(* Logix 5000 project; controller TFF vendor 1 type 14 code 107 rev 33.11; software revision 33.04; part 37 of 38 *)
(* tags used below, declared in another part *)
   Config : Configuration;   // Index Array used in configuration routines
   result : DINT[2];
   SCL : SCALE;   // Scale Instruction
   AI101Alarm : ALIAS FOR AlarmAnalog[16];
   AI104Alarm : ALIAS FOR AlarmAnalog[17];
   ControlLoop_TIC101Alarm : ALIAS FOR AlarmDeviation[7];
   FlowPath : FlowPath[64];   // Flow Path Array
   LI101 : ALIAS FOR AnalogPoint[44];
   LI101Alarm : ALIAS FOR AlarmAnalog[44];
   Options : Options;   // Options List
   PI601Alarm : ALIAS FOR AlarmAnalog[21];
   PipeAnimation : PipeAnimation;   // HMI Pipe Animation Array
   Rack_ACT350_WI101_200L : IO_Station;   // Status of ACT350 200L
   Rack_ACT350_WI101_500L : IO_Station;   // Status of ACT350 500L
   Tank : TankManagement;   // Tank Management
   TCU101Alarm : ALIAS FOR AlarmAnalog[18];
   TCU101DF : ALIAS FOR DigitalPoint[30];
   TI101Alarm : ALIAS FOR AlarmAnalog[13];
   WI101 : ALIAS FOR AnalogPoint[15];
   WI101Alarm : ALIAS FOR AlarmAnalog[15];
(* Process, continued *)

ROUTINE TankManagement   (* ladder *)
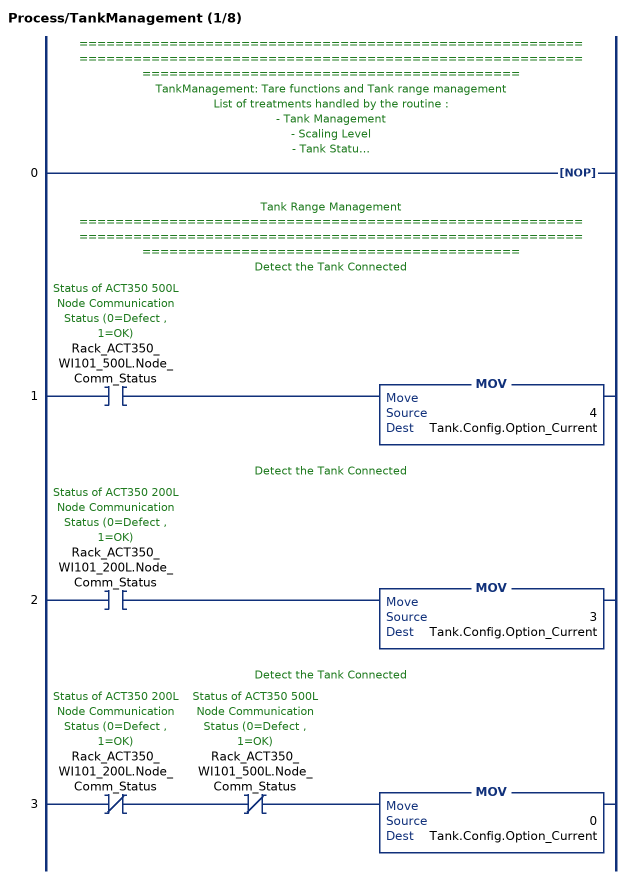
   // ==========================================================================================================================================================
   //                                                                                                                                 TankManagement: Tare functions and Tank range management
   //                                                     List of treatments handled by the routine :
   //                                                          - Tank Management
   //                                                          - Scaling Level
   //                                                          - Tank Status
   //                                                     -----------------------------------------------------------------------------------------------------------------------------------------------------
   //                                                     History
   // 		2019-DEC-24 - Merck - Q. Spindler - Initial version for Candidate Release 1.00.00.00.a
   // ==========================================================================================================================================================
   0: NOP();
   // Tank Range Management
   // ==========================================================================================================================================================
   // Detect the Tank Connected
   1: XIC(Rack_ACT350_WI101_500L.Node_Comm_Status)MOV(4,Tank.Config.Option_Current);
   // Detect the Tank Connected
   2: XIC(Rack_ACT350_WI101_200L.Node_Comm_Status)MOV(3,Tank.Config.Option_Current);
   // Detect the Tank Connected
   3: XIO(Rack_ACT350_WI101_200L.Node_Comm_Status)XIO(Rack_ACT350_WI101_500L.Node_Comm_Status)MOV(0,Tank.Config.Option_Current);
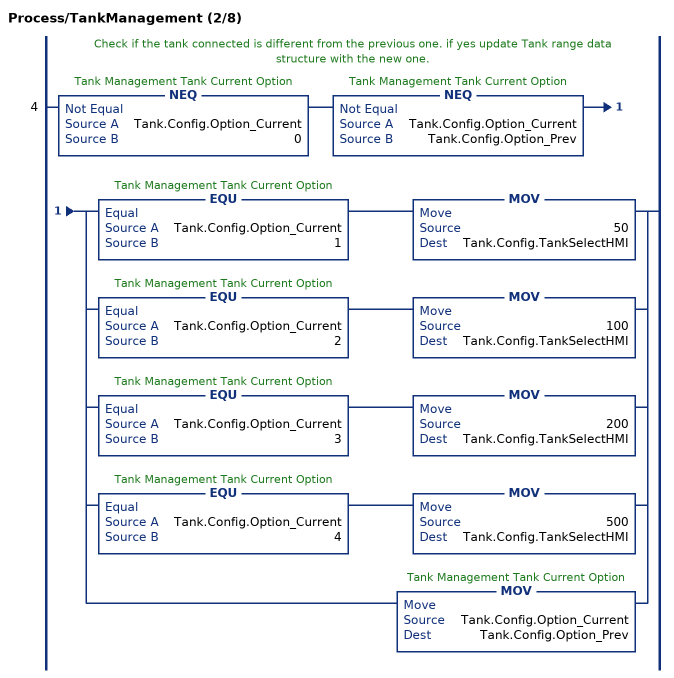
   // Check if the tank connected is different from the previous one. if yes update Tank range data structure with the new one.
   4: NEQ(Tank.Config.Option_Current,0)NEQ(Tank.Config.Option_Current,Tank.Config.Option_Prev)[[EQU(Tank.Config.Option_Current,1) MOV(50,Tank.Config.TankSelectHMI) ,EQU(Tank.Config.Option_Current,2) MOV(100,Tank.Config.TankSelectHMI) ,EQU(Tank.Config.Option_Current,3) MOV(200,Tank.Config.TankSelectHMI) ,EQU(Tank.Config.Option_Current,4) MOV(500,Tank.Config.TankSelectHMI) ] ,MOV(Tank.Config.Option_Current,Tank.Config.Option_Prev) ];
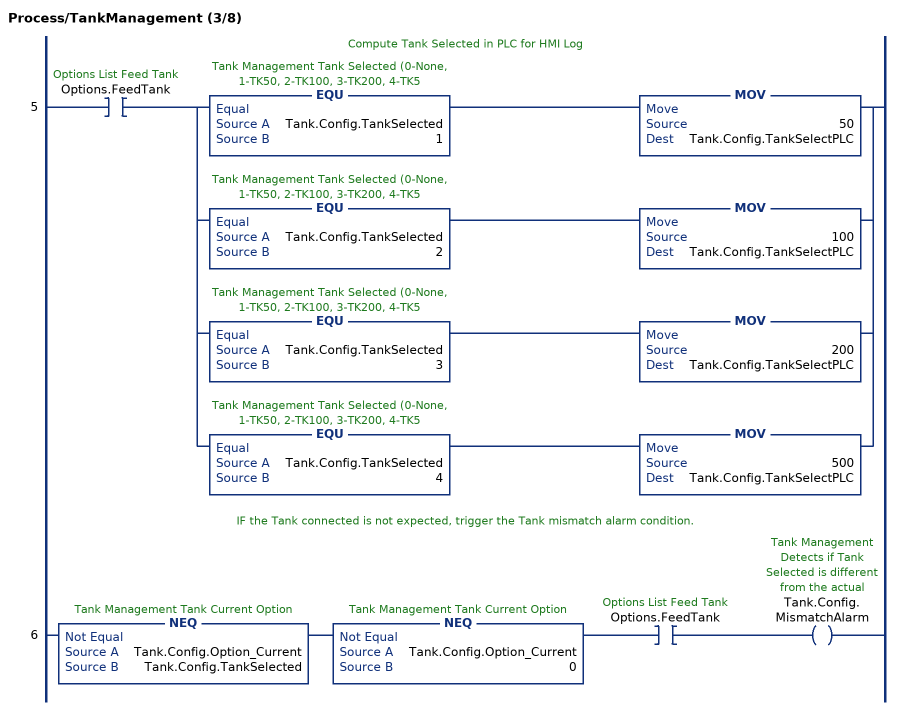
   // Compute Tank Selected in PLC for HMI Log
   5: XIC(Options.FeedTank)[EQU(Tank.Config.TankSelected,1) MOV(50,Tank.Config.TankSelectPLC) ,EQU(Tank.Config.TankSelected,2) MOV(100,Tank.Config.TankSelectPLC) ,EQU(Tank.Config.TankSelected,3) MOV(200,Tank.Config.TankSelectPLC) ,EQU(Tank.Config.TankSelected,4) MOV(500,Tank.Config.TankSelectPLC) ];
   // IF the Tank connected is not expected, trigger the Tank mismatch alarm condition.
   6: NEQ(Tank.Config.Option_Current,Tank.Config.TankSelected)NEQ(Tank.Config.Option_Current,0)XIC(Options.FeedTank)OTE(Tank.Config.MismatchAlarm);
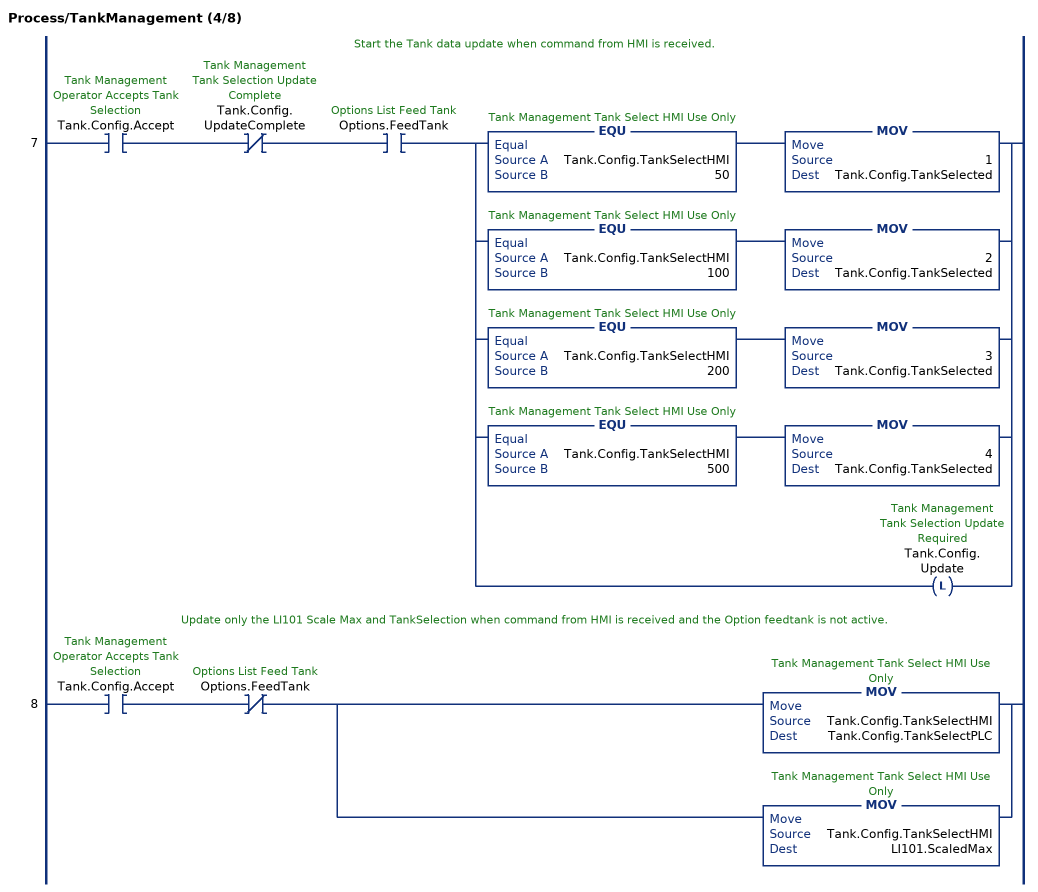
   // Start the Tank data update when command from HMI is received.
   7: XIC(Tank.Config.Accept)XIO(Tank.Config.UpdateComplete)XIC(Options.FeedTank)[[EQU(Tank.Config.TankSelectHMI,50) MOV(1,Tank.Config.TankSelected) ,EQU(Tank.Config.TankSelectHMI,100) MOV(2,Tank.Config.TankSelected) ,EQU(Tank.Config.TankSelectHMI,200) MOV(3,Tank.Config.TankSelected) ,EQU(Tank.Config.TankSelectHMI,500) MOV(4,Tank.Config.TankSelected) ] ,OTL(Tank.Config.Update) ];
   // Update only the LI101 Scale Max and TankSelection when command from HMI is received and the Option feedtank is not active.
   8: XIC(Tank.Config.Accept)XIO(Options.FeedTank)[MOV(Tank.Config.TankSelectHMI,Tank.Config.TankSelectPLC) ,MOV(Tank.Config.TankSelectHMI,LI101.ScaledMax) ];
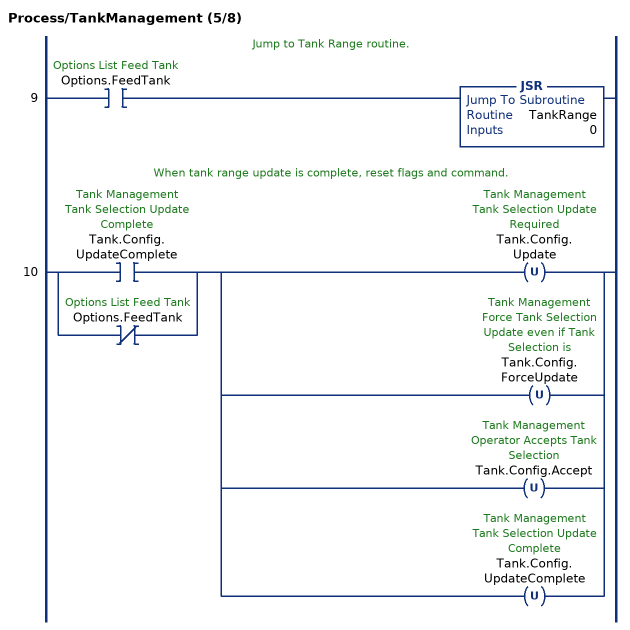
   // Jump to Tank Range routine.
   9: XIC(Options.FeedTank)JSR(TankRange,0);
   // When tank range update is complete, reset flags and command.
   10: [XIC(Tank.Config.UpdateComplete) ,XIO(Options.FeedTank) ][OTU(Tank.Config.Update) ,OTU(Tank.Config.ForceUpdate) ,OTU(Tank.Config.Accept) ,OTU(Tank.Config.UpdateComplete) ];
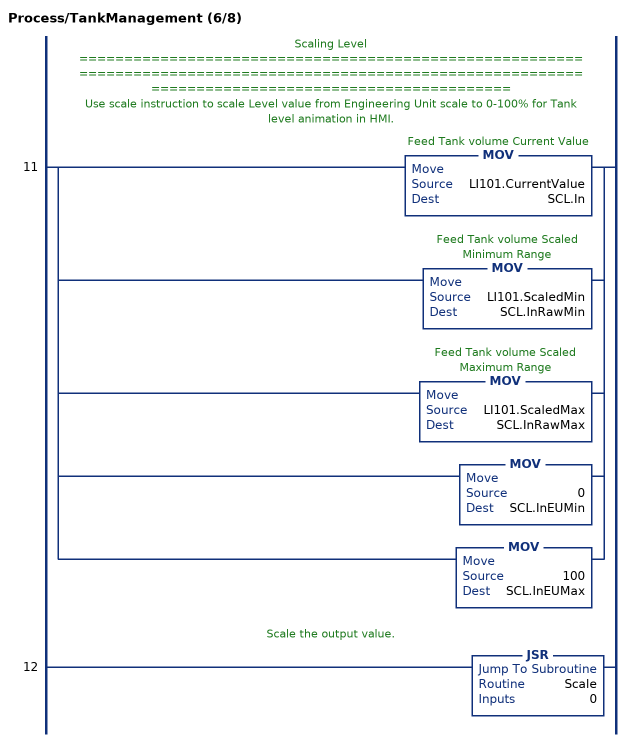
   // Scaling Level
   // ========================================================================================================================================================
   // Use scale instruction to scale Level value from Engineering Unit scale to 0-100% for Tank level animation in HMI.
   11: [MOV(LI101.CurrentValue,SCL.In) ,MOV(LI101.ScaledMin,SCL.InRawMin) ,MOV(LI101.ScaledMax,SCL.InRawMax) ,MOV(0,SCL.InEUMin) ,MOV(100,SCL.InEUMax) ];
   // Scale the output value.
   12: JSR(Scale,0);
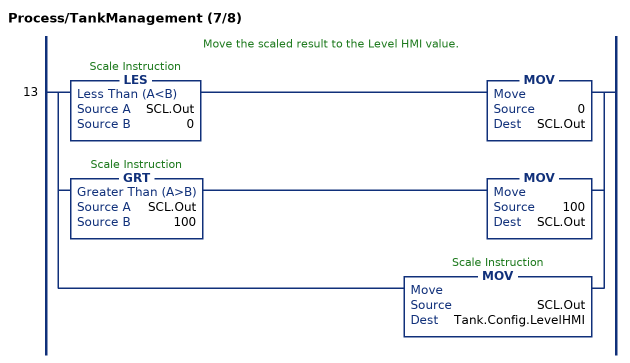
   // Move the scaled result to the Level HMI value.
   13: [LES(SCL.Out,0) MOV(0,SCL.Out) ,GRT(SCL.Out,100) MOV(100,SCL.Out) ,MOV(SCL.Out,Tank.Config.LevelHMI) ];
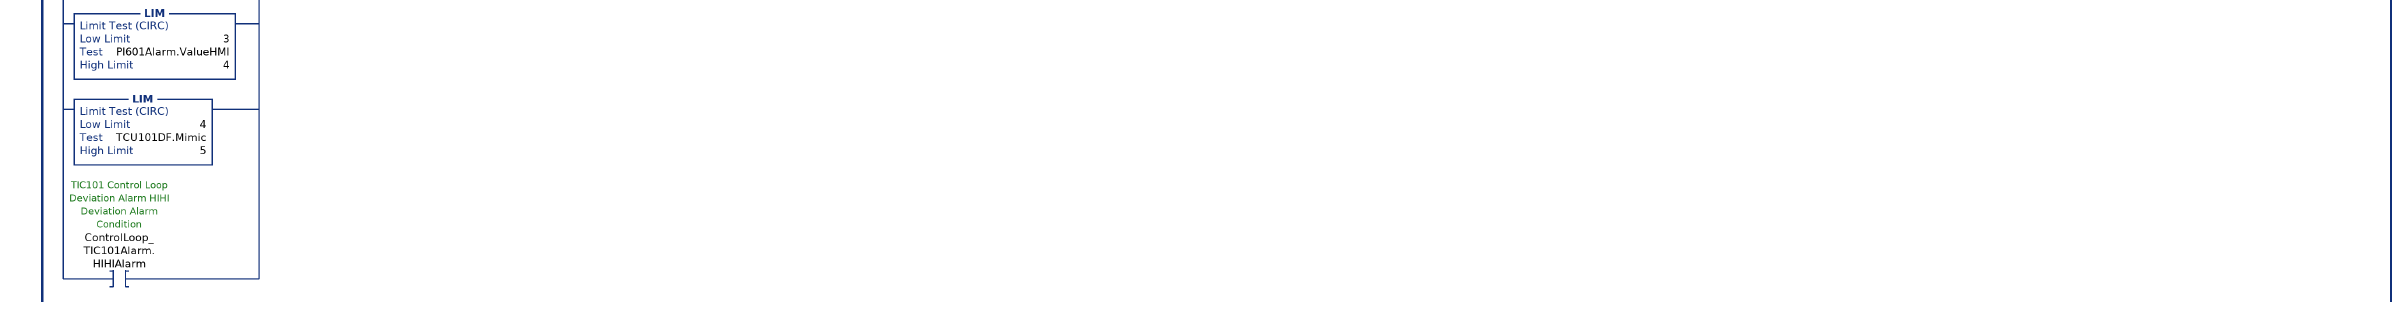
   // Tank Status
   // ==========================================================================================================================================================
   // TankAlarmStatus : 0 = No Alarm & No Flowpath Valid
   // TankAlarmStatus : 1 = No Alarm & Flowpath Valid
   // TankAlarmStatus : 2 = Tank in Non-Critical Alarm
   // TankAlarmStatus : 3 = Tank in Critical Alarm
   14: [XIO(PipeAnimation.PipeStatP1[23]) XIO(PipeAnimation.PipeStatP2[10]) LES(WI101Alarm.ValueHMI,1) LES(LI101Alarm.ValueHMI,1) LES(TI101Alarm.ValueHMI,1) LES(TCU101Alarm.ValueHMI,1) LES(AI101Alarm.ValueHMI,1) LES(AI104Alarm.ValueHMI,1) LES(PI601Alarm.ValueHMI,1) LES(TCU101DF.Mimic,2) XIO(ControlLoop_TIC101Alarm.HIAlarm) XIO(ControlLoop_TIC101Alarm.HIHIAlarm) MOV(0,Tank.Config.AlarmStatus) ,[XIC(PipeAnimation.PipeStatP1[23]) ,XIC(PipeAnimation.PipeStatP2[10]) ] LES(WI101Alarm.ValueHMI,1) LES(LI101Alarm.ValueHMI,1) LES(TI101Alarm.ValueHMI,1) LES(TCU101Alarm.ValueHMI,1) LES(AI101Alarm.ValueHMI,1) LES(AI104Alarm.ValueHMI,1) LES(PI601Alarm.ValueHMI,1) LES(TCU101DF.Mimic,2) XIO(ControlLoop_TIC101Alarm.HIAlarm) XIO(ControlLoop_TIC101Alarm.HIHIAlarm) MOV(1,Tank.Config.AlarmStatus) ,[LIM(1,WI101Alarm.ValueHMI,2) ,LIM(1,LI101Alarm.ValueHMI,2) ,LIM(1,TI101Alarm.ValueHMI,2) ,LIM(1,TCU101Alarm.ValueHMI,2) ,LIM(1,AI101Alarm.ValueHMI,2) ,LIM(1,AI104Alarm.ValueHMI,2) ,LIM(1,PI601Alarm.ValueHMI,2) ,LIM(2,TCU101DF.Mimic,3) ,XIC(ControlLoop_TIC101Alarm.HIAlarm) XIO(ControlLoop_TIC101Alarm.HIHIAlarm) ] MOV(2,Tank.Config.AlarmStatus) ,[LIM(3,WI101Alarm.ValueHMI,4) ,LIM(3,LI101Alarm.ValueHMI,4) ,LIM(3,TI101Alarm.ValueHMI,4) ,LIM(3,TCU101Alarm.ValueHMI,4) ,LIM(3,AI101Alarm.ValueHMI,4) ,LIM(3,AI104Alarm.ValueHMI,4) ,LIM(3,PI601Alarm.ValueHMI,4) ,LIM(4,TCU101DF.Mimic,5) ,XIC(ControlLoop_TIC101Alarm.HIHIAlarm) ] MOV(3,Tank.Config.AlarmStatus) ];
END_ROUTINE

ROUTINE TankRange   (* ladder *)
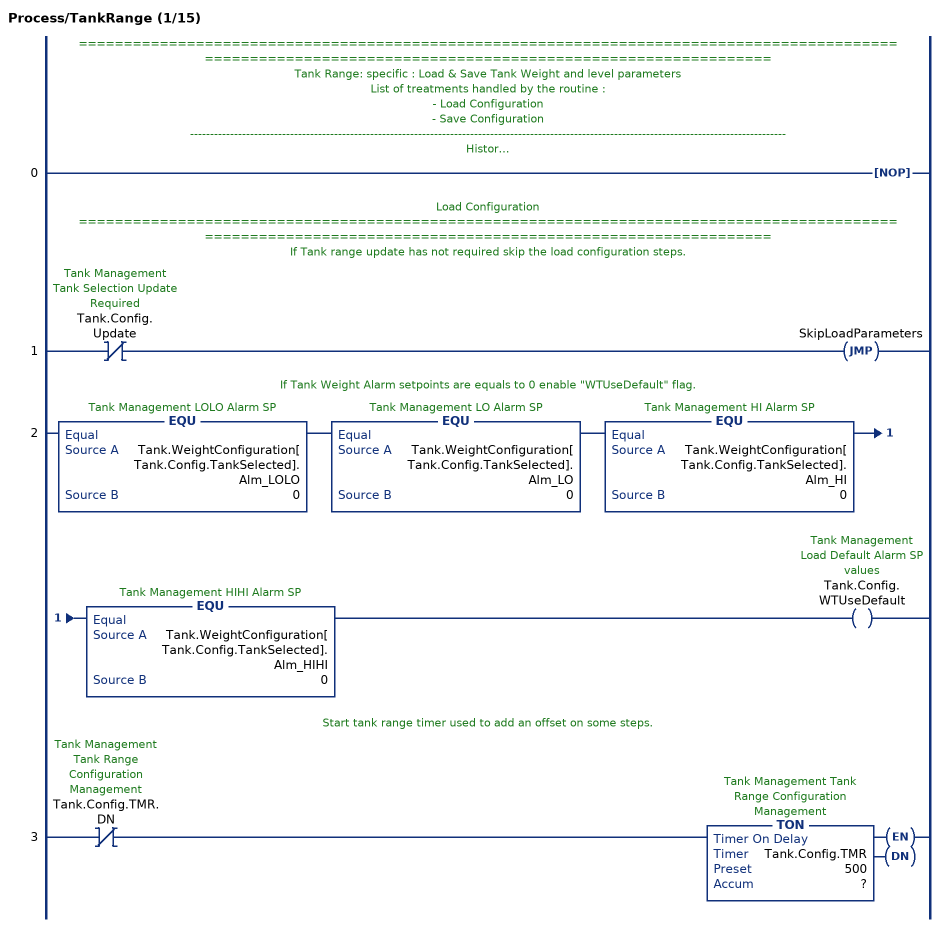
   // ==========================================================================================================================================================
   //                                                                                                                                 Tank Range: specific : Load & Save Tank Weight and level parameters
   //                                                     List of treatments handled by the routine :
   //                                                          - Load Configuration
   //                                                          - Save Configuration
   //                                                     -----------------------------------------------------------------------------------------------------------------------------------------------------
   //                                                     History
   // 		2019-DEC-24 - Merck - Q. Spindler - Initial version for Candidate Release 1.00.00.00.a
   // ==========================================================================================================================================================
   0: NOP();
   // Load Configuration
   // ==========================================================================================================================================================
   // If Tank range update has not required skip the load configuration steps.
   1: XIO(Tank.Config.Update)JMP(SkipLoadParameters);
   // If Tank Weight Alarm setpoints are equals to 0 enable "WTUseDefault" flag.
   2: EQU(Tank.WeightConfiguration[Tank.Config.TankSelected].Alm_LOLO,0)EQU(Tank.WeightConfiguration[Tank.Config.TankSelected].Alm_LO,0)EQU(Tank.WeightConfiguration[Tank.Config.TankSelected].Alm_HI,0)EQU(Tank.WeightConfiguration[Tank.Config.TankSelected].Alm_HIHI,0)OTE(Tank.Config.WTUseDefault);
   // Start tank range timer used to add an offset on some steps.
   3: XIO(Tank.Config.TMR.DN)TON(Tank.Config.TMR,?,?);
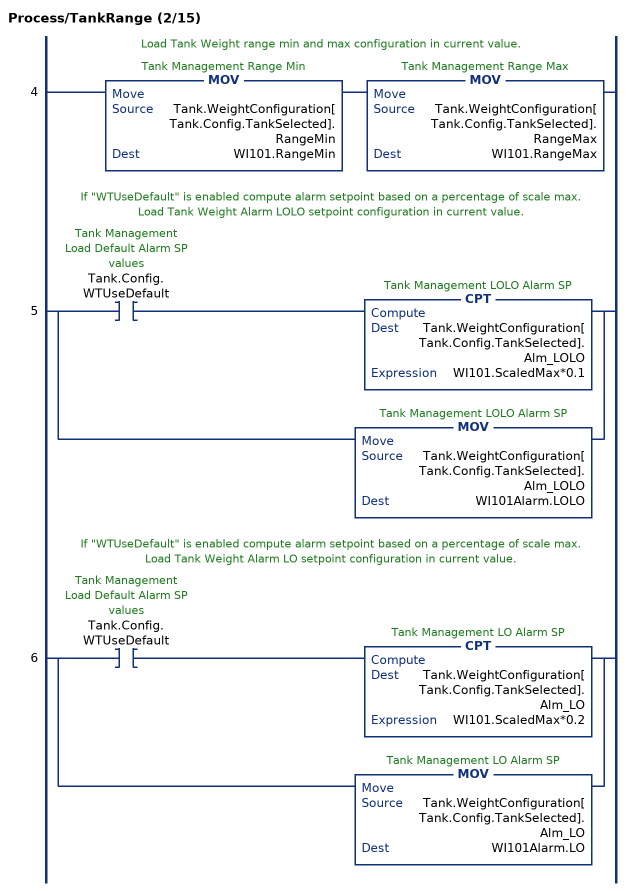
   // Load Tank Weight range min and max configuration in current value.
   4: MOV(Tank.WeightConfiguration[Tank.Config.TankSelected].RangeMin,WI101.RangeMin)MOV(Tank.WeightConfiguration[Tank.Config.TankSelected].RangeMax,WI101.RangeMax);
   // If "WTUseDefault" is enabled compute alarm setpoint based on a percentage of scale max. Load Tank Weight Alarm LOLO setpoint configuration in current value.
   5: [XIC(Tank.Config.WTUseDefault) CPT(Tank.WeightConfiguration[Tank.Config.TankSelected].Alm_LOLO,WI101.ScaledMax*0.1) ,MOV(Tank.WeightConfiguration[Tank.Config.TankSelected].Alm_LOLO,WI101Alarm.LOLO) ];
   // If "WTUseDefault" is enabled compute alarm setpoint based on a percentage of scale max. Load Tank Weight Alarm LO setpoint configuration in current value.
   6: [XIC(Tank.Config.WTUseDefault) CPT(Tank.WeightConfiguration[Tank.Config.TankSelected].Alm_LO,WI101.ScaledMax*0.2) ,MOV(Tank.WeightConfiguration[Tank.Config.TankSelected].Alm_LO,WI101Alarm.LO) ];
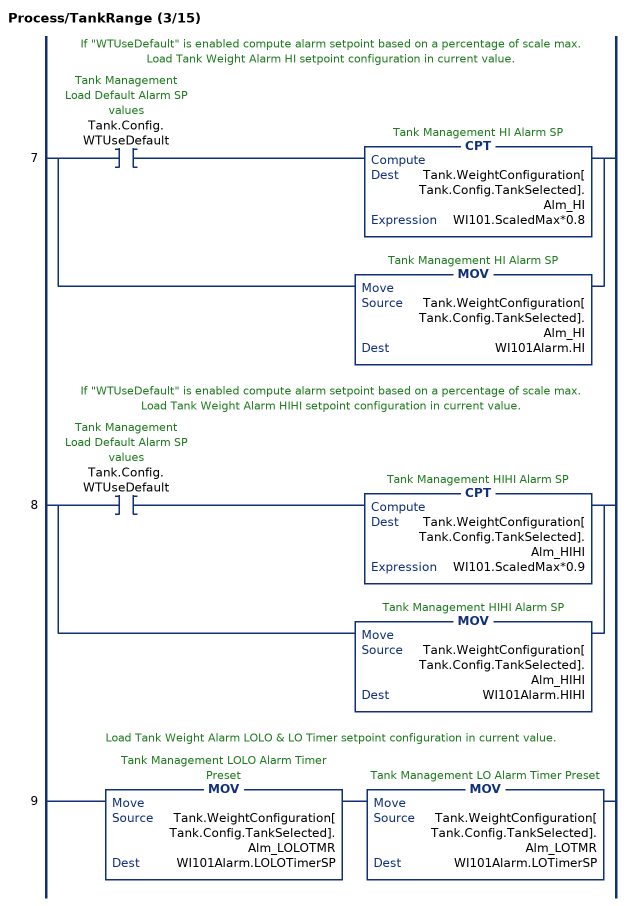
   // If "WTUseDefault" is enabled compute alarm setpoint based on a percentage of scale max. Load Tank Weight Alarm HI setpoint configuration in current value.
   7: [XIC(Tank.Config.WTUseDefault) CPT(Tank.WeightConfiguration[Tank.Config.TankSelected].Alm_HI,WI101.ScaledMax*0.8) ,MOV(Tank.WeightConfiguration[Tank.Config.TankSelected].Alm_HI,WI101Alarm.HI) ];
   // If "WTUseDefault" is enabled compute alarm setpoint based on a percentage of scale max. Load Tank Weight Alarm HIHI setpoint configuration in current value.
   8: [XIC(Tank.Config.WTUseDefault) CPT(Tank.WeightConfiguration[Tank.Config.TankSelected].Alm_HIHI,WI101.ScaledMax*0.9) ,MOV(Tank.WeightConfiguration[Tank.Config.TankSelected].Alm_HIHI,WI101Alarm.HIHI) ];
   // Load Tank Weight Alarm LOLO & LO Timer setpoint configuration in current value.
   9: MOV(Tank.WeightConfiguration[Tank.Config.TankSelected].Alm_LOLOTMR,WI101Alarm.LOLOTimerSP)MOV(Tank.WeightConfiguration[Tank.Config.TankSelected].Alm_LOTMR,WI101Alarm.LOTimerSP);
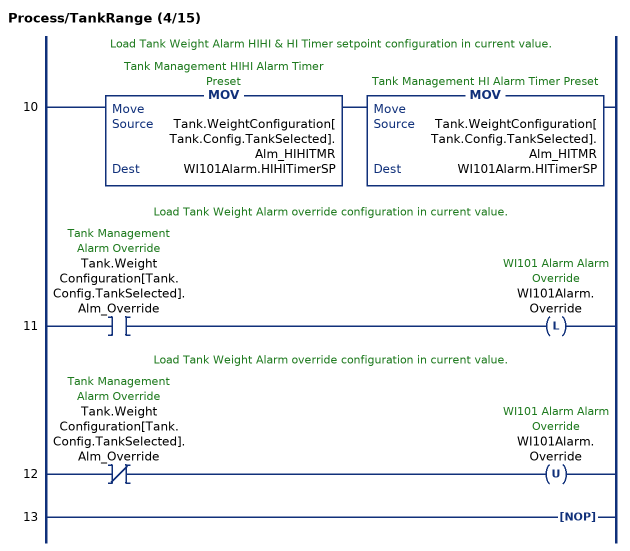
   // Load Tank Weight Alarm HIHI & HI Timer setpoint configuration in current value.
   10: MOV(Tank.WeightConfiguration[Tank.Config.TankSelected].Alm_HIHITMR,WI101Alarm.HIHITimerSP)MOV(Tank.WeightConfiguration[Tank.Config.TankSelected].Alm_HITMR,WI101Alarm.HITimerSP);
   // Load Tank Weight Alarm override configuration in current value.
   11: XIC(Tank.WeightConfiguration[Tank.Config.TankSelected].Alm_Override)OTL(WI101Alarm.Override);
   // Load Tank Weight Alarm override configuration in current value.
   12: XIO(Tank.WeightConfiguration[Tank.Config.TankSelected].Alm_Override)OTU(WI101Alarm.Override);
   13: NOP();
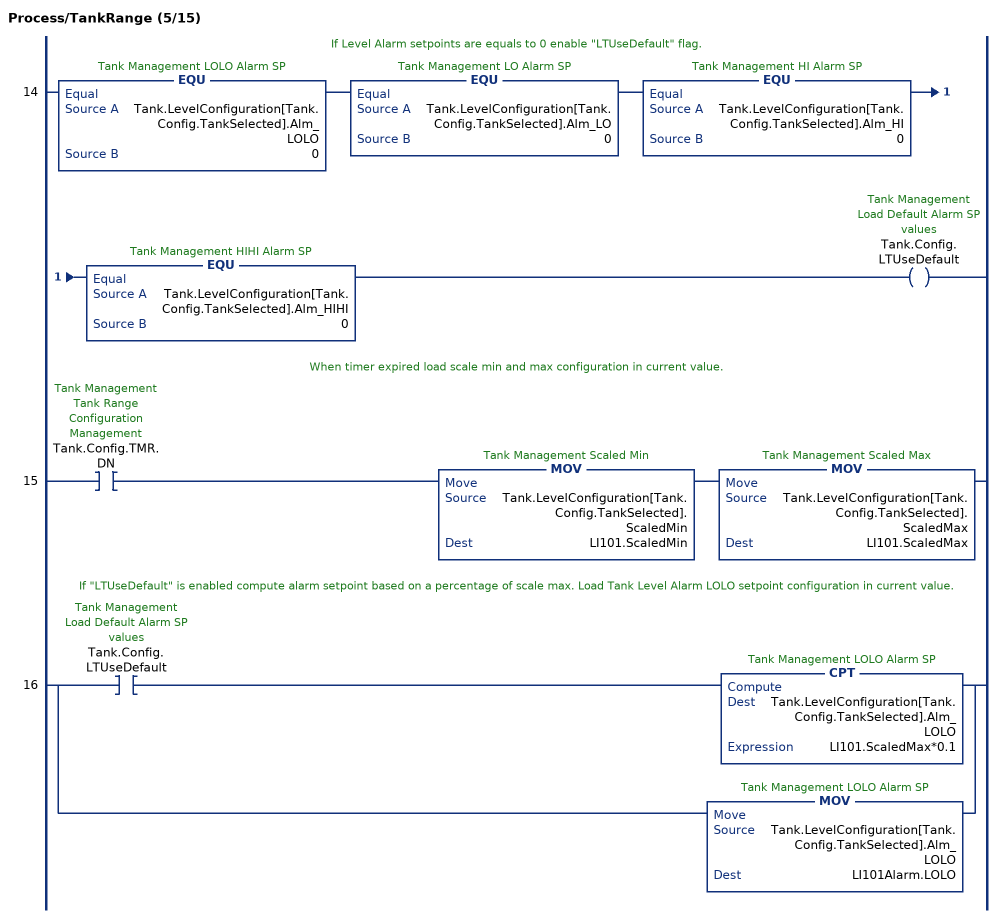
   // If Level Alarm setpoints are equals to 0 enable "LTUseDefault" flag.
   14: EQU(Tank.LevelConfiguration[Tank.Config.TankSelected].Alm_LOLO,0)EQU(Tank.LevelConfiguration[Tank.Config.TankSelected].Alm_LO,0)EQU(Tank.LevelConfiguration[Tank.Config.TankSelected].Alm_HI,0)EQU(Tank.LevelConfiguration[Tank.Config.TankSelected].Alm_HIHI,0)OTE(Tank.Config.LTUseDefault);
   // When timer expired load scale min and max configuration in current value.
   15: XIC(Tank.Config.TMR.DN)MOV(Tank.LevelConfiguration[Tank.Config.TankSelected].ScaledMin,LI101.ScaledMin)MOV(Tank.LevelConfiguration[Tank.Config.TankSelected].ScaledMax,LI101.ScaledMax);
   // If "LTUseDefault" is enabled compute alarm setpoint based on a percentage of scale max. Load Tank Level Alarm LOLO setpoint configuration in current value.
   16: [XIC(Tank.Config.LTUseDefault) CPT(Tank.LevelConfiguration[Tank.Config.TankSelected].Alm_LOLO,LI101.ScaledMax*0.1) ,MOV(Tank.LevelConfiguration[Tank.Config.TankSelected].Alm_LOLO,LI101Alarm.LOLO) ];
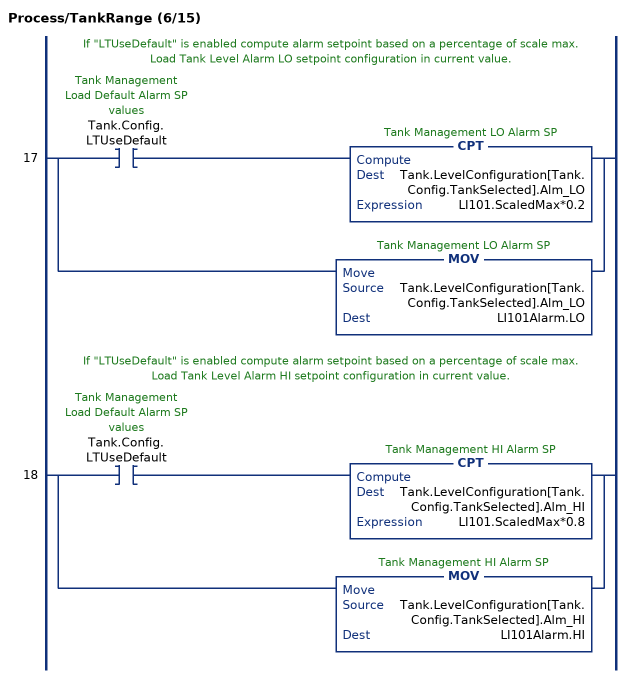
   // If "LTUseDefault" is enabled compute alarm setpoint based on a percentage of scale max. Load Tank Level Alarm LO setpoint configuration in current value.
   17: [XIC(Tank.Config.LTUseDefault) CPT(Tank.LevelConfiguration[Tank.Config.TankSelected].Alm_LO,LI101.ScaledMax*0.2) ,MOV(Tank.LevelConfiguration[Tank.Config.TankSelected].Alm_LO,LI101Alarm.LO) ];
   // If "LTUseDefault" is enabled compute alarm setpoint based on a percentage of scale max. Load Tank Level Alarm HI setpoint configuration in current value.
   18: [XIC(Tank.Config.LTUseDefault) CPT(Tank.LevelConfiguration[Tank.Config.TankSelected].Alm_HI,LI101.ScaledMax*0.8) ,MOV(Tank.LevelConfiguration[Tank.Config.TankSelected].Alm_HI,LI101Alarm.HI) ];
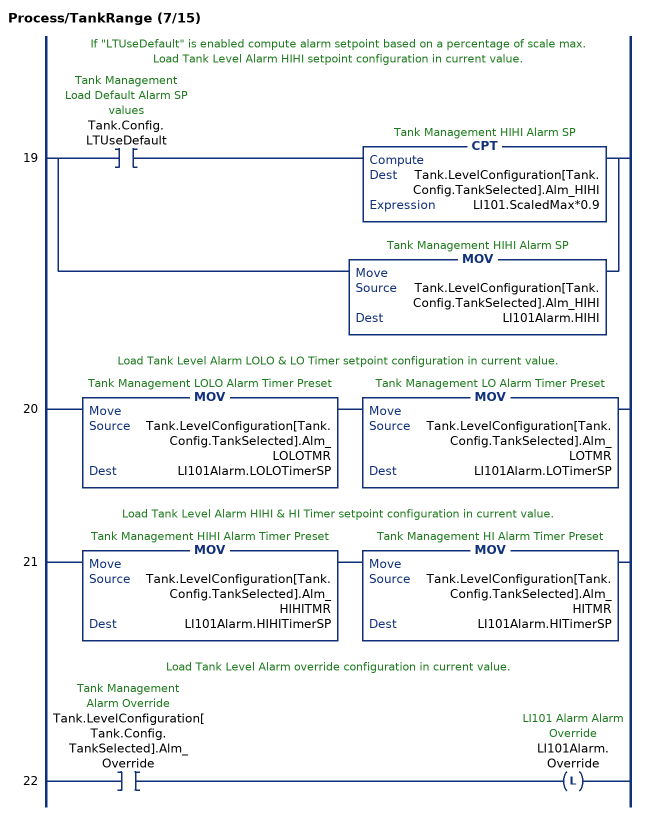
   // If "LTUseDefault" is enabled compute alarm setpoint based on a percentage of scale max. Load Tank Level Alarm HIHI setpoint configuration in current value.
   19: [XIC(Tank.Config.LTUseDefault) CPT(Tank.LevelConfiguration[Tank.Config.TankSelected].Alm_HIHI,LI101.ScaledMax*0.9) ,MOV(Tank.LevelConfiguration[Tank.Config.TankSelected].Alm_HIHI,LI101Alarm.HIHI) ];
   // Load Tank Level Alarm LOLO & LO Timer setpoint configuration in current value.
   20: MOV(Tank.LevelConfiguration[Tank.Config.TankSelected].Alm_LOLOTMR,LI101Alarm.LOLOTimerSP)MOV(Tank.LevelConfiguration[Tank.Config.TankSelected].Alm_LOTMR,LI101Alarm.LOTimerSP);
   // Load Tank Level Alarm HIHI & HI Timer setpoint configuration in current value.
   21: MOV(Tank.LevelConfiguration[Tank.Config.TankSelected].Alm_HIHITMR,LI101Alarm.HIHITimerSP)MOV(Tank.LevelConfiguration[Tank.Config.TankSelected].Alm_HITMR,LI101Alarm.HITimerSP);
   // Load Tank Level Alarm override configuration in current value.
   22: XIC(Tank.LevelConfiguration[Tank.Config.TankSelected].Alm_Override)OTL(LI101Alarm.Override);
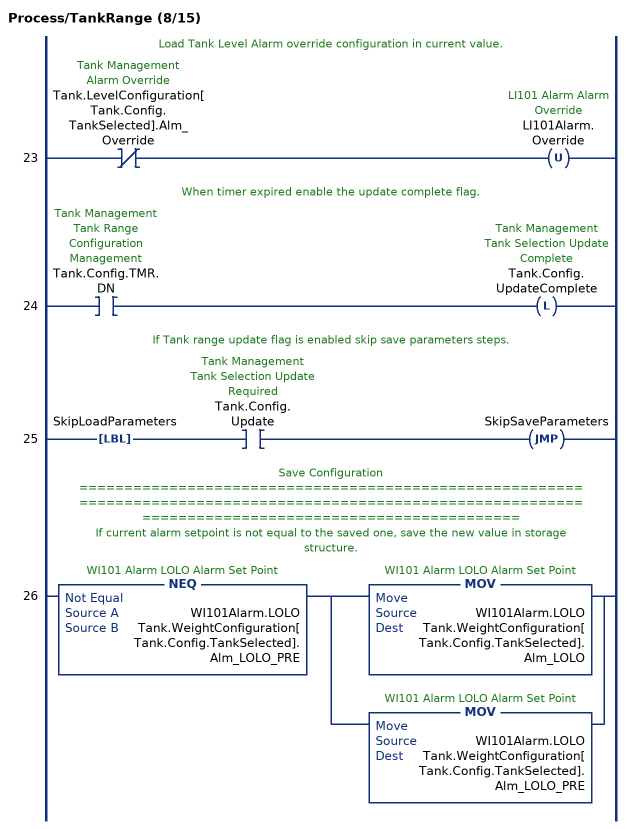
   // Load Tank Level Alarm override configuration in current value.
   23: XIO(Tank.LevelConfiguration[Tank.Config.TankSelected].Alm_Override)OTU(LI101Alarm.Override);
   // When timer expired enable the update complete flag.
   24: XIC(Tank.Config.TMR.DN)OTL(Tank.Config.UpdateComplete);
   // If Tank range update flag is enabled skip save parameters steps.
   25: LBL(SkipLoadParameters)XIC(Tank.Config.Update)JMP(SkipSaveParameters);
   // Save Configuration
   // ==========================================================================================================================================================
   // If current alarm setpoint is not equal to the saved one, save the new value in storage structure.
   26: NEQ(WI101Alarm.LOLO,Tank.WeightConfiguration[Tank.Config.TankSelected].Alm_LOLO_PRE)[MOV(WI101Alarm.LOLO,Tank.WeightConfiguration[Tank.Config.TankSelected].Alm_LOLO) ,MOV(WI101Alarm.LOLO,Tank.WeightConfiguration[Tank.Config.TankSelected].Alm_LOLO_PRE) ];
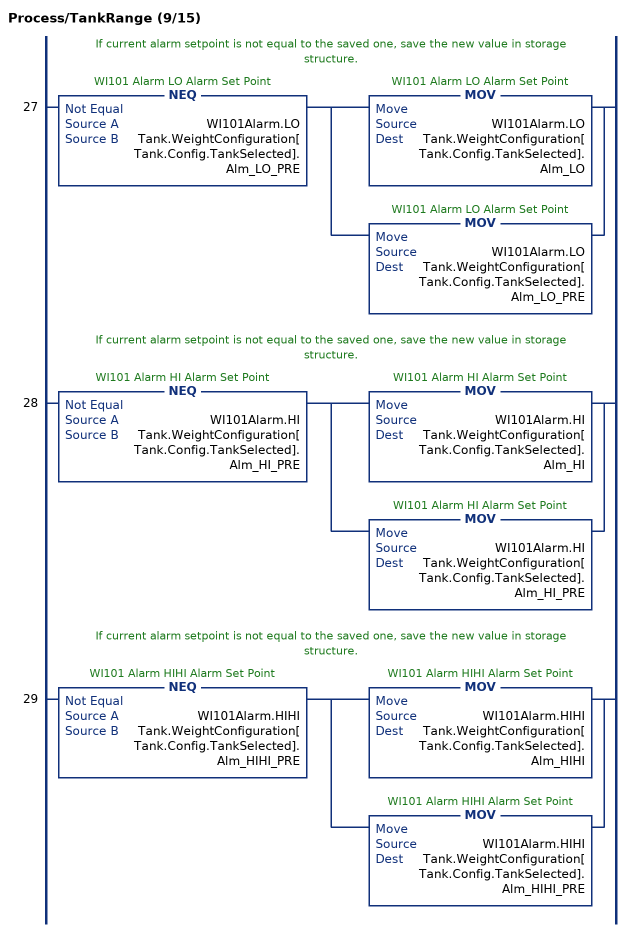
   // If current alarm setpoint is not equal to the saved one, save the new value in storage structure.
   27: NEQ(WI101Alarm.LO,Tank.WeightConfiguration[Tank.Config.TankSelected].Alm_LO_PRE)[MOV(WI101Alarm.LO,Tank.WeightConfiguration[Tank.Config.TankSelected].Alm_LO) ,MOV(WI101Alarm.LO,Tank.WeightConfiguration[Tank.Config.TankSelected].Alm_LO_PRE) ];
   // If current alarm setpoint is not equal to the saved one, save the new value in storage structure.
   28: NEQ(WI101Alarm.HI,Tank.WeightConfiguration[Tank.Config.TankSelected].Alm_HI_PRE)[MOV(WI101Alarm.HI,Tank.WeightConfiguration[Tank.Config.TankSelected].Alm_HI) ,MOV(WI101Alarm.HI,Tank.WeightConfiguration[Tank.Config.TankSelected].Alm_HI_PRE) ];
   // If current alarm setpoint is not equal to the saved one, save the new value in storage structure.
   29: NEQ(WI101Alarm.HIHI,Tank.WeightConfiguration[Tank.Config.TankSelected].Alm_HIHI_PRE)[MOV(WI101Alarm.HIHI,Tank.WeightConfiguration[Tank.Config.TankSelected].Alm_HIHI) ,MOV(WI101Alarm.HIHI,Tank.WeightConfiguration[Tank.Config.TankSelected].Alm_HIHI_PRE) ];
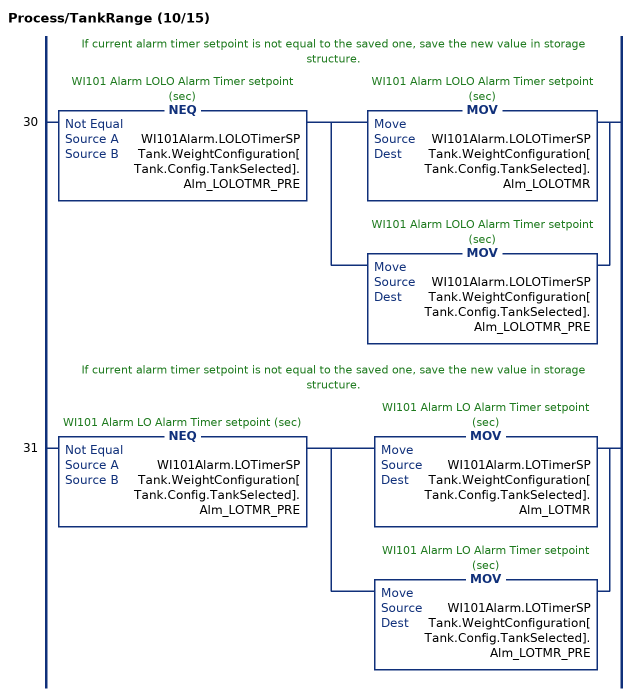
   // If current alarm timer setpoint is not equal to the saved one, save the new value in storage structure.
   30: NEQ(WI101Alarm.LOLOTimerSP,Tank.WeightConfiguration[Tank.Config.TankSelected].Alm_LOLOTMR_PRE)[MOV(WI101Alarm.LOLOTimerSP,Tank.WeightConfiguration[Tank.Config.TankSelected].Alm_LOLOTMR) ,MOV(WI101Alarm.LOLOTimerSP,Tank.WeightConfiguration[Tank.Config.TankSelected].Alm_LOLOTMR_PRE) ];
   // If current alarm timer setpoint is not equal to the saved one, save the new value in storage structure.
   31: NEQ(WI101Alarm.LOTimerSP,Tank.WeightConfiguration[Tank.Config.TankSelected].Alm_LOTMR_PRE)[MOV(WI101Alarm.LOTimerSP,Tank.WeightConfiguration[Tank.Config.TankSelected].Alm_LOTMR) ,MOV(WI101Alarm.LOTimerSP,Tank.WeightConfiguration[Tank.Config.TankSelected].Alm_LOTMR_PRE) ];
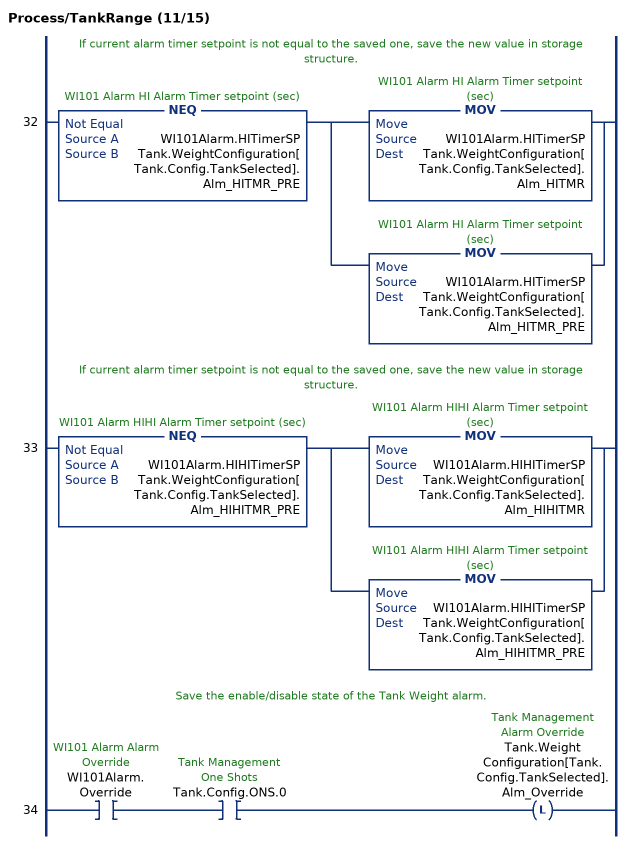
   // If current alarm timer setpoint is not equal to the saved one, save the new value in storage structure.
   32: NEQ(WI101Alarm.HITimerSP,Tank.WeightConfiguration[Tank.Config.TankSelected].Alm_HITMR_PRE)[MOV(WI101Alarm.HITimerSP,Tank.WeightConfiguration[Tank.Config.TankSelected].Alm_HITMR) ,MOV(WI101Alarm.HITimerSP,Tank.WeightConfiguration[Tank.Config.TankSelected].Alm_HITMR_PRE) ];
   // If current alarm timer setpoint is not equal to the saved one, save the new value in storage structure.
   33: NEQ(WI101Alarm.HIHITimerSP,Tank.WeightConfiguration[Tank.Config.TankSelected].Alm_HIHITMR_PRE)[MOV(WI101Alarm.HIHITimerSP,Tank.WeightConfiguration[Tank.Config.TankSelected].Alm_HIHITMR) ,MOV(WI101Alarm.HIHITimerSP,Tank.WeightConfiguration[Tank.Config.TankSelected].Alm_HIHITMR_PRE) ];
   // Save the enable/disable state of the Tank Weight alarm.
   34: XIC(WI101Alarm.Override)XIC(Tank.Config.ONS.0)OTL(Tank.WeightConfiguration[Tank.Config.TankSelected].Alm_Override);
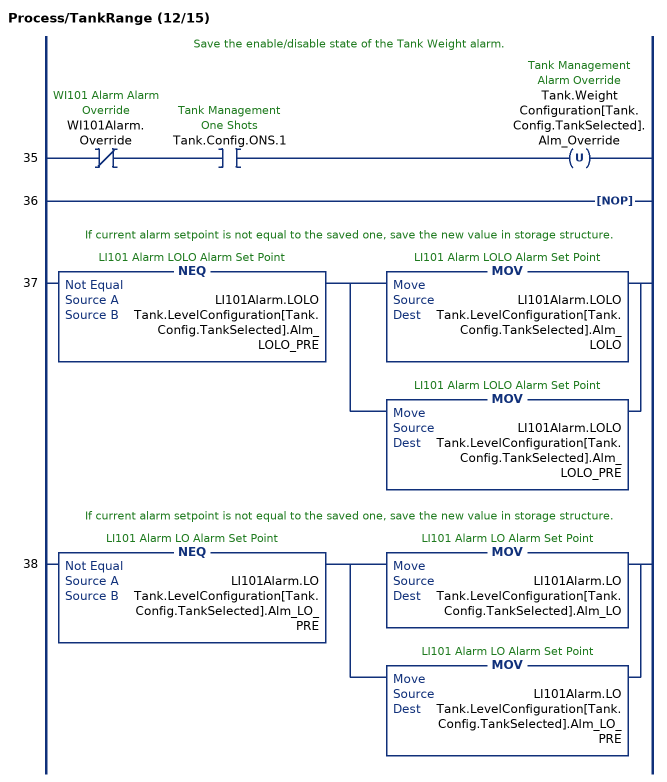
   // Save the enable/disable state of the Tank Weight alarm.
   35: XIO(WI101Alarm.Override)XIC(Tank.Config.ONS.1)OTU(Tank.WeightConfiguration[Tank.Config.TankSelected].Alm_Override);
   36: NOP();
   // If current alarm setpoint is not equal to the saved one, save the new value in storage structure.
   37: NEQ(LI101Alarm.LOLO,Tank.LevelConfiguration[Tank.Config.TankSelected].Alm_LOLO_PRE)[MOV(LI101Alarm.LOLO,Tank.LevelConfiguration[Tank.Config.TankSelected].Alm_LOLO) ,MOV(LI101Alarm.LOLO,Tank.LevelConfiguration[Tank.Config.TankSelected].Alm_LOLO_PRE) ];
   // If current alarm setpoint is not equal to the saved one, save the new value in storage structure.
   38: NEQ(LI101Alarm.LO,Tank.LevelConfiguration[Tank.Config.TankSelected].Alm_LO_PRE)[MOV(LI101Alarm.LO,Tank.LevelConfiguration[Tank.Config.TankSelected].Alm_LO) ,MOV(LI101Alarm.LO,Tank.LevelConfiguration[Tank.Config.TankSelected].Alm_LO_PRE) ];
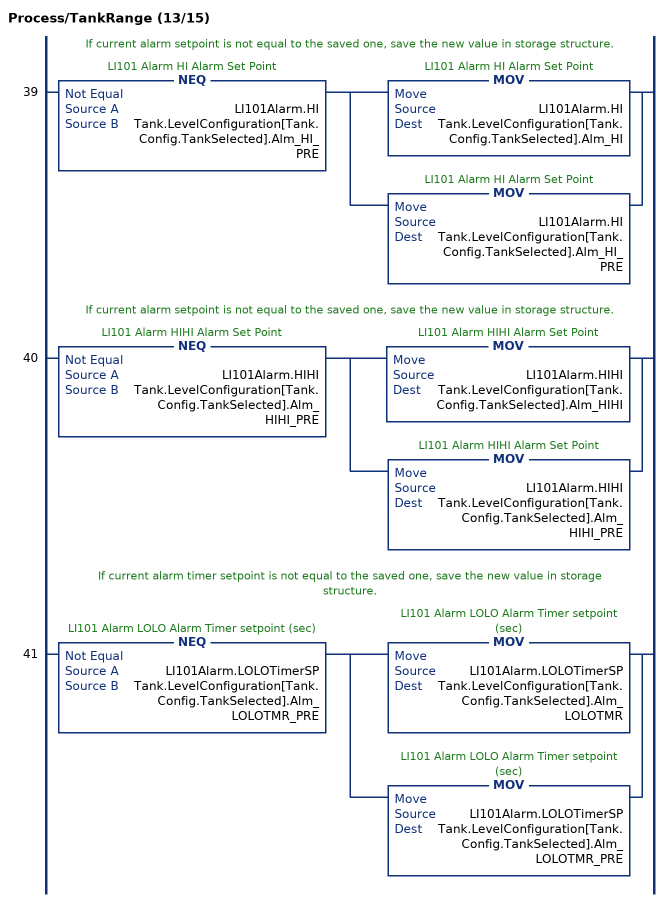
   // If current alarm setpoint is not equal to the saved one, save the new value in storage structure.
   39: NEQ(LI101Alarm.HI,Tank.LevelConfiguration[Tank.Config.TankSelected].Alm_HI_PRE)[MOV(LI101Alarm.HI,Tank.LevelConfiguration[Tank.Config.TankSelected].Alm_HI) ,MOV(LI101Alarm.HI,Tank.LevelConfiguration[Tank.Config.TankSelected].Alm_HI_PRE) ];
   // If current alarm setpoint is not equal to the saved one, save the new value in storage structure.
   40: NEQ(LI101Alarm.HIHI,Tank.LevelConfiguration[Tank.Config.TankSelected].Alm_HIHI_PRE)[MOV(LI101Alarm.HIHI,Tank.LevelConfiguration[Tank.Config.TankSelected].Alm_HIHI) ,MOV(LI101Alarm.HIHI,Tank.LevelConfiguration[Tank.Config.TankSelected].Alm_HIHI_PRE) ];
   // If current alarm timer setpoint is not equal to the saved one, save the new value in storage structure.
   41: NEQ(LI101Alarm.LOLOTimerSP,Tank.LevelConfiguration[Tank.Config.TankSelected].Alm_LOLOTMR_PRE)[MOV(LI101Alarm.LOLOTimerSP,Tank.LevelConfiguration[Tank.Config.TankSelected].Alm_LOLOTMR) ,MOV(LI101Alarm.LOLOTimerSP,Tank.LevelConfiguration[Tank.Config.TankSelected].Alm_LOLOTMR_PRE) ];
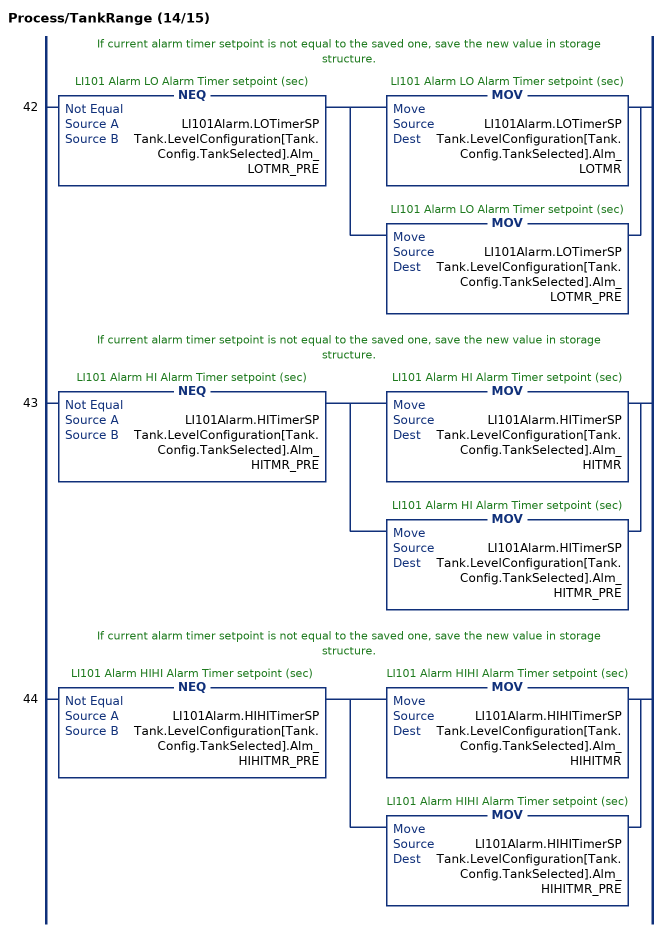
   // If current alarm timer setpoint is not equal to the saved one, save the new value in storage structure.
   42: NEQ(LI101Alarm.LOTimerSP,Tank.LevelConfiguration[Tank.Config.TankSelected].Alm_LOTMR_PRE)[MOV(LI101Alarm.LOTimerSP,Tank.LevelConfiguration[Tank.Config.TankSelected].Alm_LOTMR) ,MOV(LI101Alarm.LOTimerSP,Tank.LevelConfiguration[Tank.Config.TankSelected].Alm_LOTMR_PRE) ];
   // If current alarm timer setpoint is not equal to the saved one, save the new value in storage structure.
   43: NEQ(LI101Alarm.HITimerSP,Tank.LevelConfiguration[Tank.Config.TankSelected].Alm_HITMR_PRE)[MOV(LI101Alarm.HITimerSP,Tank.LevelConfiguration[Tank.Config.TankSelected].Alm_HITMR) ,MOV(LI101Alarm.HITimerSP,Tank.LevelConfiguration[Tank.Config.TankSelected].Alm_HITMR_PRE) ];
   // If current alarm timer setpoint is not equal to the saved one, save the new value in storage structure.
   44: NEQ(LI101Alarm.HIHITimerSP,Tank.LevelConfiguration[Tank.Config.TankSelected].Alm_HIHITMR_PRE)[MOV(LI101Alarm.HIHITimerSP,Tank.LevelConfiguration[Tank.Config.TankSelected].Alm_HIHITMR) ,MOV(LI101Alarm.HIHITimerSP,Tank.LevelConfiguration[Tank.Config.TankSelected].Alm_HIHITMR_PRE) ];
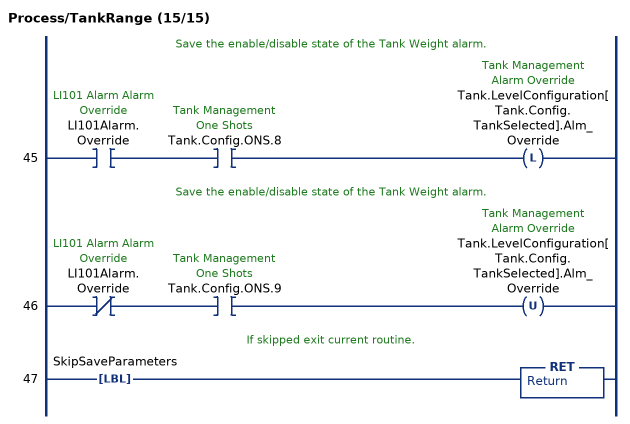
   // Save the enable/disable state of the Tank Weight alarm.
   45: XIC(LI101Alarm.Override)XIC(Tank.Config.ONS.8)OTL(Tank.LevelConfiguration[Tank.Config.TankSelected].Alm_Override);
   // Save the enable/disable state of the Tank Weight alarm.
   46: XIO(LI101Alarm.Override)XIC(Tank.Config.ONS.9)OTU(Tank.LevelConfiguration[Tank.Config.TankSelected].Alm_Override);
   // If skipped exit current routine.
   47: LBL(SkipSaveParameters)RET();
END_ROUTINE
